TYPE E_MoveMode :
(
    eAbsolute := 0,
    eRelative := 1,
    eVelocity := 2
) DINT;
END_TYPE

(* stored: Version 1.1.0.1, ProductVersion 3.1.4024.12
   DUT E_MoveMode: Id {85421ccf-6536-535e-aaa5-df51a1ac4778} *)
